FUNCTION_BLOCK ButtonM (* Composite Function Block Type *)
  (* Standard: 61499-2 *)
  (* Version 0.0, 6/20/2016, Andrei, nxtControl GmbH, template *)
  PACKAGE Main;
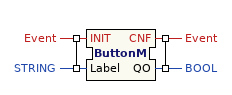
  EVENT_INPUT
    INIT WITH Label;
  END_EVENT
  EVENT_OUTPUT
    CNF WITH QO; (* Execution Confirmation *)
  END_EVENT
  VAR_INPUT
    Label : STRING;
  END_VAR
  VAR_OUTPUT
    QO : BOOL; (* Output event qualifier *)
  END_VAR
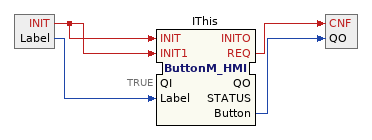
  FBS
    IThis : ButtonM_HMI(QI := TRUE);
  END_FBS
  EVENT_CONNECTIONS
    INIT TO IThis.INIT;
    IThis.REQ TO CNF;
    INIT TO IThis.INIT1;
  END_CONNECTIONS
  DATA_CONNECTIONS
    Label TO IThis.Label;
    IThis.Button TO QO;
  END_CONNECTIONS
END_FUNCTION_BLOCK
